// TIA Portal V21 export
Screen "AreaPrototypes"  1366x663
  ScreenLayer "Layer_0"
    FaceplateContainer "ManualSelector" at 245,10 size 260x34  Text="Band ein / Belt on / Band aan"
      FunctionID := 100
      Operability := Permissions.Manual
      Command := Manual.Selected
      VendorExtension 
    IOField "RecipeValue" at 245,50 size 260x34  Mode=InputOutput, Tag=Recipe.Real[0]
      OperabilityAnimation   Tag=Permissions.Parameters
    Button "Navigate" at 245,600 size 260x34
      on Press: OpenScreen(ScreenNo := 1)
    IOField "OptionalBelt" at 520,50 size 260x34  Mode=Output, Tag="Area.HMI".Belts[1].Speed
      VisibilityAnimation   RangeStart=1, RangeEnd=1, Tag="Area.HMI".Belts[1].Installed
